(* IEC 61131-3 sources: axsharp/src/sanbox/integration/ix-integration-plc/src, 12 files *)

(* ---- measurement.st ---- *)
NAMESPACE MeasurementExample
    {#ix-attr:[Container(Layout.Wrap)]}
    {#ix-attr:[Group(GroupLayout.GroupBox)]}
    {S7.extern=ReadWrite}
    CLASS PUBLIC Measurement
        VAR PUBLIC
            {#ix-set:AttributeName = "Minimum"}
            Min : REAL;
            {#ix-set:AttributeName = "Measured"}
            {#ix-attr:[ReadOnly()]}
            Acquired : REAL;
            {#ix-set:AttributeName = "Maximum"}
            Max : REAL;
            {#ix-set:AttributeName = "Measurement Result"}
            Result : Result;
        END_VAR

        METHOD PUBLIC Simulate
            Min := Min - REAL#1.0;
            Max := Max + REAL#1.0;
            Max := Max / REAL#2.0;
        END_METHOD
    END_CLASS

    TYPE
        Result : INT (
            None := 0,
            Passed := 10,
            Failed := 20
        );
    END_TYPE

    {S7.extern=ReadWrite}
    CLASS PUBLIC Measurements
        VAR PUBLIC
            {#ix-attr:[Container(Layout.Stack)]}
            {#ix-attr:[Group(GroupLayout.GroupBox)]}
            {#ix-set:AttributeName = "Stack panel"}
            measurement_stack : Measurement;

            {#ix-attr:[Container(Layout.Wrap)]}
            {#ix-attr:[Group(GroupLayout.GroupBox)]}
            {#ix-set:AttributeName = "Wrap panel"}
            measurement_wrap : Measurement;

            {#ix-attr:[Container(Layout.UniformGrid)]}
            {#ix-attr:[Group(GroupLayout.GroupBox)]}
            {#ix-set:AttributeName = "Grid"}
            measurement_grid : Measurement;

            {#ix-attr:[Container(Layout.Tabs)]}
            {#ix-attr:[Group(GroupLayout.GroupBox)]}
            {#ix-set:AttributeName = "Tabs"}
            measurement_tabs : Measurement;
        END_VAR

        METHOD PUBLIC Simulate
            measurement_stack.Simulate();
            measurement_wrap.Simulate();
            measurement_grid.Simulate();
            measurement_tabs.Simulate();
        END_METHOD

    END_CLASS
END_NAMESPACE

(* ---- weather.st ---- *)
{#ix[Container(Layout.Tabs)]}
{S7.extern=ReadWrite}
CLASS weather
    VAR PUBLIC
        GeoLocation : GeoLocation;
        {#ix[Container(Layout.Wrap)]}
        Temperature : REAL;
        Humidity : REAL;
        Location : STRING;
        ChillFactor : REAL;
        Feeling : Feeling;
    END_VAR
END_CLASS

{S7.extern=ReadWrite}
CLASS weathers
    VAR PUBLIC
        i : ARRAY[0..50] OF weatherBase;
    END_VAR
END_CLASS

TYPE
    Feeling : (Freezing, Cold, Lookworm, Warm, Hot);
END_TYPE

TYPE
    {S7.extern=ReadWrite}
    Colors : INT (
        RED := 12,
        GREEN := 14,
        BLUE := 23
    );
END_TYPE

(* ---- all_primitives.st ---- *)
USING System.Strings;

{S7.extern=ReadWrite}

CLASS all_primitives
    VAR PUBLIC
        myBOOL	        :       BOOL	      ;
        myBYTE	        :       BYTE	      := BYTE#1;
        myWORD	        :       WORD	      := WORD#1;
        myDWORD	        :       DWORD	      := DWORD#1;
        myLWORD	        :       LWORD	      := LWORD#1;
        mySINT	        :       SINT	      ;
        myINT	        :       INT	          ;
        myDINT	        :       DINT	      ;
        myLINT	        :       LINT	      ;
        myUSINT	        :       USINT	      ;
        myUINT	        :       UINT	      ;
        myUDINT	        :       UDINT	      ;
        myULINT	        :       ULINT	      ;
        myREAL	        :       REAL	      ;
        myLREAL	        :       LREAL	      ;
        myTIME	        :       TIME	      ;
        myLTIME	        :       LTIME	      ;
        myDATE	        :       DATE	      ;
        myLDATE	        :       LDATE	      ;
        myTIME_OF_DAY	:       TIME_OF_DAY	  ;
        myLTIME_OF_DAY	:       LTIME_OF_DAY  ;
        myDATE_AND_TIME  :      DATE_AND_TIME ;
        myLDATE_AND_TIME :      LDATE_AND_TIME;
        myCHAR	        :       CHAR	      ;
        myWCHAR	        :       WCHAR	      ;
        mySTRING	        :   STRING	      ;
        myWSTRING	    :       WSTRING	      ;

        testLWORD : LWORD;
        testULINT : ULINT;
        testULINTPlusOne : ULINT;
        testLWORDPlusOne : LWORD;

    END_VAR

    METHOD PUBLIC Simulate

      myBOOL := NOT myBOOL;
      myBYTE := TO_BYTE(TO_SINT(myBYTE) + 1);
      myWORD := TO_WORD(TO_INT(myWORD) + 1);
      myDWORD := TO_DWORD(TO_DINT(myDWORD) + 1);
      myLWORD := TO_LWORD(TO_LINT(myLWORD) + 1);
      mySINT := mySINT + SINT#1;
      myINT := myINT + 1;
      myDINT := myDINT + DINT#1;
      myLINT := myLINT + LINT#1;
      myUSINT := myUSINT + USINT#1;
      myUINT := myUINT + UINT#1;
      myUDINT := myUDINT + UDINT#1;
      myULINT := myULINT + ULINT#1;
      myREAL := myREAL + REAL#1.0;
      myLREAL := myLREAL + 1.0;
      myTIME := myTIME + T#1s;
      myLTIME := myLTIME + LT#1s;
      myDATE := TO_DATE(To_LWORD(TO_ULINT(TO_LWORD(myDATE)) + ULINT#86400000000000));
      myLDATE := TO_DATE(To_LWORD(TO_ULINT(TO_LWORD(myLDATE)) + ULINT#86400000000000));
      myTIME_OF_DAY := myTIME_OF_DAY + T#1s;
      myLTIME_OF_DAY := myLTIME_OF_DAY + LT#1s;
      myDATE_AND_TIME := myDATE_AND_TIME + T#1s;
      myLDATE_AND_TIME := myLDATE_AND_TIME + LT#1s;
      myCHAR := myCHAR + CHAR#1;
      myWCHAR := myWCHAR + WCHAR#1;
      mySTRING := ToString(myINT);
      //myWSTRING := ToString(myINT);
  END_METHOD
END_CLASS

(* ---- compositeLayout.st ---- *)
{S7.extern=ReadWrite}
CLASS compositeLayout
    VAR PUBLIC
        {#ix-set:AttributeName = "<#Integer From PLC#>"}
        testInteger : INT;
        {#ix-set:AttributeName = "<#UInteger From PLC#>"}
        testUInteger : INT;
        {#ix-set:AttributeName = "<#STRING From PLC#>"}
        testString : STRING;
        {#ix-set:AttributeName = "<#Task#>"}
        myTask: taskExample;
        testReal : REAL;
        {#ix-set:AttributeName = "<#LREAL From PLC#>"}
        testLReal : LREAL;
        {#ix-set:AttributeName = "<#BOOL From PLC#>"}
        testBool : BOOL;
        {#ix-set:AttributeName = "<#DATE From PLC#>"}
        TestDate : DATE;
        {#ix-set:AttributeName = "<#DATE_AND_TIME From PLC#>"}
        TestDateTime : DATE_AND_TIME;
        {#ix-set:AttributeName = "<#TIME_OF_DAY From PLC#>"}
        TestTimeOfDay : TIME_OF_DAY;
    END_VAR

END_CLASS

(* ---- example.st ---- *)
{S7.extern=ReadWrite}
CLASS example
    VAR PUBLIC
        {#ix-attr:[Container(Layout.Stack)]}
        primitives_stack: test_primitive;
        {#ix-attr:[Container(Layout.Wrap)]}
        primitives_wrap: test_primitive;
        {#ix-attr:[Container(Layout.Tabs)]}
        primitives_tabs: test_primitive;
        {#ix-attr:[Container(Layout.UniformGrid)]}
        primitives_uniform: test_primitive;

        {#ix-attr:[Container(Layout.Stack)]}
        {#ix-attr:[Group(GroupLayout.GroupBox)]}
        test_groupbox: test_primitive;

        {#ix-attr:[Container(Layout.Stack)]}
        {#ix-attr:[Group(GroupLayout.Border)]}
        test_border: test_primitive;

        {#ix-attr:[Container(Layout.Tabs)]}
        {#ix-attr:[Group(GroupLayout.GroupBox)]}
        testgroupbox: groupbox;
        testborder: border;

        ixcomponent_instance: ixcomponent;
        ixcomponent_instance2: MySecondNamespace.ixcomponent;
        ixcomponent_instance3: ThirdNamespace.ixcomponent;

        {#ix-attr:[Container(Layout.Stack)]}
        compositeStack :compositeLayout;
        {#ix-attr:[Container(Layout.Wrap)]}
        compositeWrap :compositeLayout;
        {#ix-attr:[Container(Layout.UniformGrid)]}
        compositeUniform :compositeLayout;
        {#ix-attr:[Container(Layout.Tabs)]}
        compositeTabs :compositeLayout;

        refIxComponent : REF_TO ixcomponent;
    END_VAR

    METHOD PUBLIC ReferenceToComponent : Int
        refIxComponent^ := ixcomponent_instance;
    END_METHOD

END_CLASS

(* ---- geolocation.st ---- *)
{#ix-attr:[Container(Layout.Stack)]}
{#ix-attr:[Group(GroupLayout.GroupBox)]}
{#ix-set:AttributeName = "Location"}
{S7.extern=ReadWrite}
CLASS  GeoLocation
    VAR PUBLIC
        {#ix-set:AttributeName = "Latitude [°]"}
        {#ix-set:AttributeMinimum = -90.0f}
        {#ix-set:AttributeMaximum = 90.0f}
        Latitude : REAL;
        {#ix-set:AttributeName = "Logitude [°]"}
        {#ix-set:AttributeMinimum = 0.0f}
        {#ix-set:AttributeMaximum = 180.0f}
        Longitude : REAL;
        {#ix-set:AttributeName = "Altitude [m]"}
        Altitude : REAL;
        {#ix-set:AttributeName = "Short descriptor"}
        Description : STRING[10];
        {#ix-set:AttributeName = "Long descriptor"}
        LongDescription : STRING[254];
    END_VAR
END_CLASS

(* ---- ixcomponent.st ---- *)
{S7.extern=ReadWrite}
CLASS ixcomponent
    VAR PUBLIC
        {#ix-set:AttributeName = "My integer"}
        my_int : INT;
        {#ix-set:AttributeName = "My string"}
        my_string : STRING;
        {#ix-set:AttributeName = "My bool"}
        my_bool : BOOL;
    END_VAR

    METHOD PUBLIC Simulate
        my_int := my_int + INT#1;
    END_METHOD
END_CLASS

NAMESPACE MySecondNamespace
    {S7.extern=ReadWrite}
    CLASS ixcomponent
        VAR PUBLIC
            {#ix-set:AttributeName = "My integer"}
            my_int : INT;
            {#ix-set:AttributeName = "My string"}
            my_string : STRING;
            {#ix-set:AttributeName = "My bool"}
            my_bool : BOOL;
        END_VAR
    END_CLASS
END_NAMESPACE

NAMESPACE ThirdNamespace
    {S7.extern=ReadWrite}
    CLASS ixcomponent
        VAR PUBLIC
            {#ix-set:AttributeName = "My integer"}
            my_int : INT;
            {#ix-set:AttributeName = "My string"}
            my_string : STRING;
            {#ix-set:AttributeName = "My bool"}
            my_bool : BOOL;
        END_VAR
    END_CLASS
END_NAMESPACE

(* ---- monster.st ---- *)
NAMESPACE MonsterData
    {S7.extern=ReadWrite}
    CLASS MonsterBase
        VAR PUBLIC
            ArrayOfBytes : ARRAY[0..3] OF BYTE;
            ArrayOfDrives : ARRAY[0..3] OF DriveBase;
            ArrayOfIxComponent : ARRAY[0..3] OF ixcomponent;
        END_VAR
    END_CLASS

    {S7.extern=ReadWrite}
    CLASS Monster EXTENDS MonsterBase
        VAR PUBLIC
            DriveA : DriveBase;
        END_VAR
    END_CLASS

    {S7.extern=ReadWrite}
    CLASS DriveBase
        VAR PUBLIC
            Position : LREAL;
            Velo : LREAL;
            Acc : LREAL;
            Dcc : LREAL;
        END_VAR
    END_CLASS
END_NAMESPACE

(* ---- taskExample.st ---- *)
{S7.extern=ReadWrite}
CLASS TaskExample
    VAR PUBLIC
        example : STRING;
    END_VAR

END_CLASS

(* ---- weatherBase.st ---- *)
    {#ix-attr:[Container(Layout.Stack)]}
    {#ix-attr:[Group(GroupLayout.GroupBox)]}
    {S7.extern=ReadWrite}
    CLASS PUBLIC weatherBase
      VAR PUBLIC
        Latitude : REAL;
        Longitude : REAL;
        Altitude : REAL;
        Description : STRING;
        {#ix-attr:[ReadOnly()]}
        LongDescription : STRING;
        {#ix-attr:[ReadOnce()]}
        {#ix-set:AttributeName = "this has [ReadOnce()] attribute will be readon only once..."}
        StartCounter : INT;

        {#ix-attr:[RenderIgnore()]}
        {#ix-set:AttributeName = "[RenderIgnore()] must not be displayed!"}
        RenderIgnoreAllToghether : STRING;
        {#ix-set:AttributeName = "[RenderIgnore(''Control'')]"}
        {#ix-attr:[RenderIgnore("Control")]}
        RenderIgnoreWhenControl : STRING;
        {#ix-set:AttributeName = "[RenderIgnore(''Display'')]"}
        {#ix-attr:[RenderIgnore("Display")]}
        RenderIgnoreWhenDisplay : STRING;
        {#ix-set:AttributeName = "[RenderIgnore(''Control'', ''ShadowControl'')]"}
        {#ix-attr:[RenderIgnore("Control", "ShadowControl")]}
        RenderIgnoreWhenControlAndShadow : STRING;
        {#ix-set:AttributeName = "[RenderIgnore(''Display'', ''ShadowDisplay'')]"}
        {#ix-attr:[RenderIgnore("Display", "ShadowDisplay")]}
        RenderIgnoreWhenDisplayAndShadow : STRING;
      END_VAR
    END_CLASS

(* ---- configuration.st ---- *)
USING MonsterData;
CONFIGURATION MyConfiguration
    TASK Main(Interval := T#10ms, Priority := 1);
    PROGRAM P1 WITH Main: MyProgram;

    VAR_GLOBAL
        {S7.extern=ReadWrite}
        all_primitives : all_primitives;
        {S7.extern=ReadWrite}
        weather : weather;
        {S7.extern=ReadWrite}
        weathers : weathers;
        {S7.extern=ReadWrite}
        {#ix-set:AttributeName = "Weather in a stack pannel and grouped in group box"}
        weather_stacked : Layouts.Stacked.weather;
        {S7.extern=ReadWrite}
        {#ix-set:AttributeName = "Weather in a wrap pannel and grouped in group box"}
        weather_wrapped : Layouts.Wrapped.weather;
        {S7.extern=ReadWrite}
        {#ix-set:AttributeName = "Weather in a tabs and grouped in group box"}
        weather_tabbed : Layouts.Tabbed.weather;
        {S7.extern=ReadWrite}
        {#ix-set:AttributeName = "Weather structure set to read once"}
        {#ix-attr:[ReadOnce()]}
        weather_readOnce : Layouts.Stacked.weather;
        {S7.extern=ReadWrite}
        {#ix-set:AttributeName = "Weather structure set to read only"}
        {#ix-attr:[ReadOnly()]}
        {S7.extern=ReadWrite}
        weather_readOnly : Layouts.Stacked.weather;

        {S7.extern=ReadWrite}
        test_example: example;
        {S7.extern=ReadWrite}
        measurements : MeasurementExample.Measurements;
        {S7.extern=ReadWrite}
        ixcomponent : ixcomponent;
        {S7.extern=ReadWrite}
        monster : Monster;

        {S7.extern=ReadWrite}
        test_all_primitives : all_primitives;
    END_VAR
END_CONFIGURATION

(* ---- program.st ---- *)
PROGRAM MyProgram
    VAR_EXTERNAL
        all_primitives : all_primitives;
        weather_stacked : Layouts.Stacked.weather;
        weather_wrapped : Layouts.Wrapped.weather;
        weather_tabbed : Layouts.Tabbed.weather;
        weather_readOnce : Layouts.Stacked.weather;
        test_example: example;
        measurements : MeasurementExample.Measurements;
        ixcomponent : ixcomponent;

        test_all_primitives : all_primitives;
    END_VAR

    VAR

    END_VAR

    VAR_TEMP

    END_VAR
    all_primitives.myINT := all_primitives.myINT + 1;
    weather_stacked.Altitude := all_primitives.myINT;
    weather_wrapped.Altitude := all_primitives.myINT;
    weather_tabbed.Altitude := all_primitives.myINT;
    weather_readOnce.Altitude := all_primitives.myINT;

    weather_stacked.StartCounter := all_primitives.myINT;
    weather_wrapped.StartCounter := all_primitives.myINT;
    weather_tabbed.StartCounter := all_primitives.myINT;
    weather_readOnce.StartCounter := all_primitives.myINT;

    measurements.Simulate();
    ixcomponent.Simulate();

    test_all_primitives.Simulate();

END_PROGRAM
